Universal Robots PolyScope program: external_control.urp

Program external_control (installation=ursim_docker directory=/ursim/programs createdIn=5.26.1 lastSavedIn=5.26.1 robotSerialNumber=20195599999)
Calibrated DH parameters: a=[0, -0.425, -0.3922, 0, 0, 0]; d=[0.1625, 0, 0, 0.1333, 0.0997, 0.0996]; alpha=[1.570796, 0, 0, 1.570796, -1.570796, 0]; deltaTheta=[0, 0, 0, 0, 0, 0]
InitVariablesNode
Robot Program (runOnlyOnce=false)
  MoveJ speed 60 deg/s, acceleration 80 deg/s^2 (useActiveTCP=true optimoveEnabled=false optiMoveSpeed=0.3 optiMoveAcceleration=0.09) feature=Base
    Waypoint Waypoint_1: TCP in base x=0 y=-232.9 z=1079.4 mm, rx=0 ry=2.2214 rz=-2.2214 rad; joints [0, -90, 0, -90, 0, 0] deg
  URCap External Control (External Control, FZI Research Center for Information Technology)
